FUNCTION F_TimeHhmm : UINT		// 현지 시각 → HHMM (예: 13시 5분 = 1305)
VAR_INPUT
	i_stTime	: ST_LocalTime;
END_VAR

F_TimeHhmm := i_stTime.nHour * 100 + i_stTime.nMinute;

END_FUNCTION

(* stored: Version 1.1.0.1, ProductVersion 3.1.4024.15
   POU F_TimeHhmm: Id {ccf8cc59-7ff6-4f0a-8a1a-e1857acc2a99}, SpecialFunc None *)
